Fanuc KAREL source: KA00120.KL

PROGRAM KA00120
%NOLOCKGROUP
VAR
  SRC: CONFIG
  DST: ARRAY[2] OF SHORT
BEGIN
  SRC.CFG_FLIP = TRUE
  DST[1] = SRC
END KA00120
